FUNCTION_BLOCK FB_CommandSelector
VAR_INPUT
	bManualMode : BOOL;
    bManualForward : BOOL;
    bManualBackward : BOOL;
    bAutoForward : BOOL;
    bAutoBackward : BOOL;
END_VAR

VAR_OUTPUT
	bRequestedForward : BOOL;
    bRequestedBackward : BOOL;
END_VAR

VAR
	
END_VAR

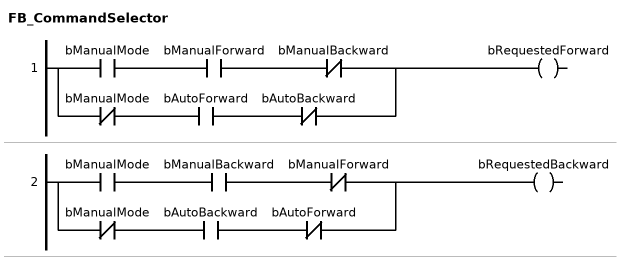
// NETWORK 1
bRequestedForward := bManualMode AND bManualForward AND NOT bManualBackward OR NOT bManualMode AND bAutoForward AND NOT bAutoBackward;

// NETWORK 2
bRequestedBackward := bManualMode AND bManualBackward AND NOT bManualForward OR NOT bManualMode AND bAutoBackward AND NOT bAutoForward;

END_FUNCTION_BLOCK

(* stored: Version 1.1.0.1
   POU FB_CommandSelector: Id {7e67a37c-c4f4-486f-b0af-c2c0600af04c}, SpecialFunc None *)
